      | 		#sleep(1.0)
      | 	#end
      | 	sleep(1.0)
      | 	#sleep(vibration_time)
      | 
      | 	movel(tilted_pose_in_base, a=0.03, v=0.1)
      | 	set_analog_out(0, 0.0)
      | 
      | 	tilt_pose_rel = pose_trans(pose_inv(p_center), tilted_pose_in_base)
      | 
      | 	lifted_pose_rel = pose_trans(lift_offset, tilt_pose_rel)
      | 
      | 	global lifted_pose = pose_trans(p_center, lifted_pose_rel)
      | 	movel(lifted_pose, a=0.03, v=0.1)
      | 	CCW_Rotate()
      | end
      | 
      | 
      | # calculate center pose on top of the container using pose transformation
      | def center_pose():
      | 	# pose transformation from side of the container to top to get center point
      | 	trans_rel = p[-0.005, 0.05, -0.027, 0, 0, 0]
      | 
      | 	p_translated = pose_trans(place_pose, trans_rel)
      | 	cx = p_translated[0]
      | 	cy = p_translated[1]
      | 	cz = p_translated[2]
      | 
      | 	global p_center_vertical = p[cx,cy,cz, 0, 0, 4.14]
      | 
      | 	#movej(p_center_vertical, a =0.3, v =0.3)
      | 	return p_center_vertical
      | end
      | 
      | # update center pose based on tilting
      | def updated_center_pose(p_center_vertical, angle_deg):
      | 	hinge_pose = pose_trans(p_center_vertical, p[0,0,-0.2,0,0,0])
      | 	local_rel = pose_trans(pose_inv(hinge_pose), p_center_vertical)
      | 
      | 	rot_tilt = p[0,0,0, -deg2rad(angle_deg),0,0]
      | 	local_rel_tilted = pose_trans(rot_tilt, local_rel)
      | 
      | 	global p_center = pose_trans(hinge_pose, local_rel_tilted)
      | 	return p_center
      | end
      | 
      | #------
      | # POTS commands
      | def tilt_send(angle):
      | 	socket_open("192.168.12.101", 80)
      | 	angle = 92.0 - angle
      | 	socket_send_string("Tilt,"+to_str(angle)+",0")
      | 	sync()
      | 	sleep(0.5)
      | 	socket_close()
      | end
      | 
      | def Motors_off():
      | 	socket_open("192.168.12.101", 80)
      | 	socket_send_string("Off,0,0")
      | 	sync()
      | 	sleep(0.5)
      | 	socket_close()
      | end
      | 
      | def Rotate():
      | 	socket_open("192.168.12.101", 80)
      | 	socket_send_string("FullRotation, 1, 2000")
      | 	sync()
      | 	sleep(0.5)
      | 	socket_close()
      | end
      | 
      | 
      | def CCW_Rotate():
      | 	socket_open("192.168.12.101", 80)
      | 	socket_send_string("FullRotation, -1, 2000")
      | 	sync()
      | 	sleep(0.5)
      | 	socket_close()
      | end
      | 
      | def tilt_to_home():
      | 	socket_open("192.168.12.101", 80)
      | 	socket_send_string("Home,0,0")
      | 	sync()
      | 	sleep(0.5)
      | 	socket_close()
      | end
    SuppressedNode
      Script file /programs/04 Scripts/dosing.script
        | def vibration_2():
        | 	set_analog_out(0,0.4)
        | 	sleep(0.8)
        | 	set_analog_out(0,0.0)
        | 	sleep(0.2)
        | end
        | 
        | def vibration_3():
        | 	set_analog_out(0,0.4)
        | 	sleep(0.5)
        | 	set_analog_out(0,0.0)
        | 	sleep(0.3)
        | end
        | 
        | def vibration_4():
        | 	set_analog_out(0,0.4)
        | 	sleep(0.6)
        | 	set_analog_out(0, 0.0)
        | 	sleep(0.5)
        | end
        | 
        | def vibration_1():
        | 	set_analog_out(0,0.4)
        | 	sleep(1)
        | 	set_analog_out(0,0.0)
        | 	sleep(0)
        | end
        | 
        | def move_tilt_in_steps(Pow_center, final_pose, steps):
        | 	i = 0
        | 	while i <= steps:
        | 		ratio = i / steps
        | 		pose_step = p[Pow_center[0] + ratio * (final_pose[0] - Pow_center[0]), Pow_center[1] + ratio * (final_pose[1] -Pow_center[1]),Pow_center[2] + ratio * (final_pose[2] - Pow_center[2]), Pow_center[3] + ratio * (final_pose[3] - Pow_center[3]), Pow_center[4] + ratio * (final_pose[4] - Pow_center[4]), Pow_center[5] + ratio * (final_pose[5] - Pow_center[5])]
        | 		movej(pose_step, a=1.2, v=0.15)
        | 		sleep(0.1)
        | 		i = i+1
        | 	end
        | end
        | 
        | def tilt_container(angle):
        | 	p_center = get_actual_tcp_pose()
        | 	hinge_offset = p[0,0,-0.23,0,0,0]
        | 	pivot_pose = pose_trans(p_center, hinge_offset)
        | 	pose_rel = pose_trans(pose_inv(pivot_pose), p_center)
        | 	angle_mid = (angle/2.0)*3.1416/180
        | 	angle_end = angle*3.1416/180
        | 	tilt_mid = p[0,0,0, -angle_mid, 0, 0]
        | 	tilt_end = p[0,0,0, -angle_end, 0, 0]
        | 	pose_rel_mid = pose_trans(tilt_mid, pose_rel)
        | 	pose_rel_end = pose_trans(tilt_end, pose_rel)
        | 	via_pose = pose_trans(pivot_pose, pose_rel_mid)
        | 	end_pose = pose_trans(pivot_pose, pose_rel_end)
        | 	movec(via_pose, end_pose, a=0.05, v=0.01, r=0.001)
        | 	p_center = get_actual_tcp_pose()
        | end
        | 
        | def deg2rad(d):
        | 	return d*3.141592/180
        | end
        | 
        | def map_tilt_to_ry_deg(container_deg):
        | 	#ry_deg = -0.875*container_deg +87.0
        | 	#return clamp(ry_deg, 5.0, 80.0)
        | 	if (Pow_name == "NaCl" or Pow_name == "Mannitol" or Pow_name == "CCS" or Pow_name == "MCC"):
        | 		if ( level>=10.0):
        | 			ry_min = 10.0
        | 			ry_max = 75.0
        | 		elif (level<10.00 and level >1.00):
        | 			ry_min = 16.0
        | 			ry_max = 65.0
        | 		else:
        | 			ry_min=17.0
        | 			ry_max=75.0
        | 		end
        | 	else:
        | 		if ( level>=10.0):
        | 			ry_min = 0.0
        | 			ry_max = 65.0
        | 		elif (level<10.00 and level >1.00):
        | 			ry_min = 10.0
        | 			ry_max = 45.0
        | 		else:
        | 			ry_min=0.0
        | 			ry_max=50.0
        | 		end
        | 
        | 	end
        | 	local span_count = angle_max -angle_min
        | 	local span_ry = ry_max - ry_min
        | 
        | 	local t = (container_deg -angle_min)/span_count
        | 	local ry_deg = ry_max - t*span_ry
        | 
        | 	return clamp(ry_deg, ry_min, ry_max)
        | 
        | end
        | 
        | def caluclate_corrections(level):
        | 	z_high = 0.01
        | 	z_low = -0.08
        | 	y_high = -0.01
        | 	y_low = -0.015
        | 
        | 	scale = (level - 10.0) / (100.0-10.0)
        | 
        | 	global correction_z = z_low + scale*(z_high - z_low)
        | 	global correction_y = y_low + scale*(y_high -y_low)
        | 
        | end
        | 
        | def scoop_powder(p_center):
        | 	#lift_offset = p[0, 0, 0.05, 0, 0, 0]
        | 	vibration_voltage = 0.4
        | 	vibration_time = 3.0
        | 	diameter = 0.07
        | 	global scoop_radius_default = 0.0
        | 	#p_center = center_pose_t
        | 
        | 
        | 	if (level >=70.00):
        | 		approach_offset = p[0.008,0,0.22,0,0,0]
        | 		lift_offset = p[0, 0, 0.05, 0, 0, 0]
        | 		caluclate_corrections(level)
        | 	elif (level >=10.00 and level <70):
        | 		approach_offset = p[0.008,0,0.22,0,0,0]
        | 		lift_offset = p[0, 0, 0.15, 0, 0, 0]
        | 		caluclate_corrections(level)
        | 	elif (level<10.00 and level >= 1.00):
        | 		approach_offset = p[0.01,0,0.22,0,0,0]
        | 		correction_z = -0.08
        | 		correction_y = -0.01
        | 		lift_offset = p[0, 0, 0.14, 0, 0, 0]
        | 	else:
        | 		approach_offset = p[0.008,0,0.22,0,0,0]
        | 		correction_z = -0.08
        | 		correction_y = -0.01
        | 		lift_offset = p[0, 0, 0.14, 0, 0, 0]
        |  	end
        | 
        | 	if (spatula == "spatula_L"):
        | 		global spatula_depth = 0.015
        | 	elif (spatula == "spatula_M"):
        | 		global spatula_depth = 0.01
        | 	elif (spatula == "spatula_S"):
        | 		global spatula_depth = 0.008
        | 	elif (spatula == "spatula_flat_M"):
        | 		global spatula_depth = 0.001
        | 	elif (spatula == "spatula_flat_S"):
        | 		global spatula_depth = 0.005
        | 	end
        | 
        | 	scoop_radius_default = diameter/2 - spatula_depth
        | 	scoop_entry_pose = pose_trans(p_center, approach_offset)
        | 	movel(scoop_entry_pose, a=0.1, v=0.25)
        | 
        | 	scoop_start_rel = p[scoop_radius_default, 0, scoop_depth, 0, 0, 0]
        | 
        | 	rot_mid = p[0, 0, 0, 0, 0, 0.785]
        | 	rot_end = p[0, 0, 0, 0, 0, 1.5708]
        | 
        | 	scoop_via_rel = pose_trans(rot_mid, scoop_start_rel)
        | 	scoop_end_rel = pose_trans(rot_end, scoop_start_rel)
        | 
        | 	scoop_start_pose = pose_trans(p_center, scoop_start_rel)
        | 	scoop_via_pose = pose_trans(p_center, scoop_via_rel)
        | 	scoop_end_pose = pose_trans(p_center, scoop_end_rel)
        | 
        | 	movel(scoop_start_pose, a=0.5, v=0.3)
        | 	#movel(p_center, a=0.5, v=1.0)
        | 	#sleep(5.0)
        | 
        | 	if (level<90.0):
        | 		Rotate()
        | 	end
        | 
        | 	#movec(scoop_via_pose, scoop_end_pose, a=0.03, v=0.05)
        | 	movec(scoop_via_pose, scoop_end_pose, a=0.03, v=0.02)
        | 	#movel(pose_trans(get_actual_tcp_pose(), p[0,0,0,0,0,deg2rad(90.0)]), a=0.03, v=0.05)
        | 	sleep(1.0)
        | 	local ry_deg = map_tilt_to_ry_deg(angle_deg)
        | 	local ry = deg2rad(ry_deg)
        | 	local end_rel = pose_trans(pose_inv(p_center), scoop_end_pose)
        | 	local end_rel_tilted = pose_trans(end_rel, p[0, 0, 0, 0, ry, 0])
        | 	global tilted_pose_in_base = pose_trans(p_center, p[0,correction_y,correction_z,end_rel_tilted[3],end_rel_tilted[4], end_rel_tilted[5]])
        | 	global tilted_pose_in_base = pose_trans(tilted_pose_in_base, p[0, 0, spatula_len, 0, 0, 0])
        | 
        | 	if (Pow_name == "lactose_fine" or Pow_name == "Magnesium_sterate"):
        | 		tilt_send((angle_deg+5))
        | 	end
        | 	movel(tilted_pose_in_base, a=0.03, v=0.1)
        | 
        | 	if (Pow_name == "lactose_fine" or Pow_name == "Magnesium_sterate"):
        | 		tilt_send((angle_deg-5))
        | 	end
        | 
        | 	if (spatula=="spatula_flat_S" or spatula=="spatula_S"):
        | 		vibration_3()
        | 	else:
        | 		set_analog_out(0, vibration_voltage)
        | 	end
        | 	if (Pow_name=="Mannitol" or Pow_name =="NaCl"):
        | 		local n=1.4
        | 	else:
        | 		local n=1.5
        | 	end
        | 	local ry_level = deg2rad(ry_deg/n)
        | 	local end_rel_tilted_level = pose_trans(end_rel, p[0, 0, 0, 0, ry_level, 0])
        | 	local level_tilted_pose_in_base = pose_trans(p_center, p[0,correction_y,correction_z,end_rel_tilted_level[3],end_rel_tilted_level[4], end_rel_tilted_level[5]])
        | 	local level_tilted_pose_in_base = pose_trans(level_tilted_pose_in_base, p[0, 0, spatula_len, 0, 0, 0])
        | 
        | 	movel(level_tilted_pose_in_base, a=0.03, v=0.1)
        | 	#if (level>70.0):
        | 		#sleep(1.0)
        | 	#end
        | 	sleep(1.0)
        | 	#sleep(vibration_time)
        | 
        | 	movel(tilted_pose_in_base, a=0.03, v=0.1)
        | 	set_analog_out(0, 0.0)
        | 
        | 	tilt_pose_rel = pose_trans(pose_inv(p_center), tilted_pose_in_base)
        | 
        | 	lifted_pose_rel = pose_trans(lift_offset, tilt_pose_rel)
        | 
        | 	global lifted_pose = pose_trans(p_center, lifted_pose_rel)
        | 	movel(lifted_pose, a=0.03, v=0.1)
        | 	CCW_Rotate()
        | end
        | 
        | 
        | def center_pose():
        | 	trans_rel = p[-0.005, 0.05, -0.015, 0, 0, 0]
        | 
        | 	p_translated = pose_trans(place_pose, trans_rel)
        | 	cx = p_translated[0]
        | 	cy = p_translated[1]
        | 	cz = p_translated[2]
        | 
        | 	global p_center_vertical = p[cx,cy,cz, 0, 0, 4.09]
        | 
        | 	#movej(p_center_vertical, a =0.3, v =0.3)
        | 	return p_center_vertical
        | end
        | 
        | def updated_center_pose(p_center_vertical, angle_deg):
        | 	hinge_pose = pose_trans(p_center_vertical, p[0,0,-0.2,0,0,0])
        | 	local_rel = pose_trans(pose_inv(hinge_pose), p_center_vertical)
        | 
        | 	rot_tilt = p[0,0,0, -deg2rad(angle_deg),0,0]
        | 	local_rel_tilted = pose_trans(rot_tilt, local_rel)
        | 
        | 	global p_center = pose_trans(hinge_pose, local_rel_tilted)
        | 	return p_center
        | end
        | 
        | def tilt_send(angle):
        | 	socket_open("192.168.12.101", 80)
        | 	angle = 92.0 - angle
        | 	socket_send_string("Tilt,"+to_str(angle)+",0")
        | 	sync()
        | 	sleep(0.5)
        | 	socket_close()
        | end
        | 
        | def Motors_off():
        | 	socket_open("192.168.12.101", 80)
        | 	socket_send_string("Off,0,0")
        | 	sync()
        | 	sleep(0.5)
        | 	socket_close()
        | end
        | 
        | def Rotate():
        | 	socket_open("192.168.12.101", 80)
        | 	socket_send_string("FullRotation, 1, 2000")
        | 	sync()
        | 	sleep(0.5)
        | 	socket_close()
        | end
        | 
        | 
        | def CCW_Rotate():
        | 	socket_open("192.168.12.101", 80)
        | 	socket_send_string("FullRotation, -1, 2000")
        | 	sync()
        | 	sleep(0.5)
        | 	socket_close()
        | end
        | def tilt_to_home():
        | 	socket_open("192.168.12.101", 80)
        | 	socket_send_string("Home,0,0")
        | 	sync()
        | 	sleep(0.5)
        | 	socket_close()
        | end
    Script file /programs/04 Scripts/Weight_scale_socket_s.script
      | def get_weight():
      | 	socket_open("192.168.12.111", 3002)
      | 	sleep(0.2)
      | 	textmsg("socket opened successfully!")
      | 	socket_send_string("GET_WEIGHT")
      | 	sync()
      | 	sleep(0.5)
      | 	receiveFromServ = socket_read_ascii_float(6)
      | 	while (receiveFromServ[0] <1):
      | 		sleep(0.5)
      | 		receiveFromServ = socket_read_ascii_float(1)
      | 		textmsg("retrying read:", receiveFromServ)
      | 	end
      | 	textmsg("Received weight:", receiveFromServ[1])
      | 	socket_close()
      | 	sleep(0.2)
      | 	return receiveFromServ[1]
      | end
      | 
      | def tare_scale():
      | 	socket_open("192.168.12.111", 3002)
      | 	socket_send_string("TARE")
      | 	sleep(0.5)
      | 	socket_close()
      | end
      | 
      | def zero_scale():
      | 	socket_open("192.168.12.111", 3002)
      | 	socket_send_string("ZERO")
      | 	sleep(0.5)
      | 	socket_close()
      | end
      | 
      | def log_weight():
      | 	socket_open("192.168.12.111", 3002)
      | 	socket_send_string("LOG_WEIGHT")
      | 	sleep(0.5)
      | 	socket_close()
      | end
      | 
      | def send_target_info():
      | 	socket_open("192.168.12.111", 3002)
      | 	socket_send_string("SET_TARGET:" + to_str(target_weight))
      | 	sleep(0.2)
      | 	socket_close()
      | end
      | def send_powder_info():
      | 	socket_open("192.168.12.111", 3002)
      | 	socket_send_string("SET_POWDER:" + Pow_name)
      | 	sleep(0.2)
      | 	socket_close()
      | end
      | def send_spatula_info():
      | 	socket_open("192.168.12.111", 3002)
      | 	socket_send_string("SET_SPATULA:" + spatula)
      | 	sleep(0.2)
      | 	socket_close()
      | end
      | 
      | def send_level_info():
      | 	socket_open("192.168.12.111",3002)
      | 	socket_send_string("SET_LEVEL:" + to_str(level))
      | 	sleep(0.2)
      | 	socket_close()
      | end
    SuppressedNode
      Script file /programs/04 Scripts/Calibration_s.script
        | # ------------------------------------------------------------
        | # Theoretical W_FULL from Cylinder Volume + Density
        | # (Eliminates manual W_FULL; keeps W_EMPTY + W_now for level)
        | # ------------------------------------------------------------
        | # -------------------------
        | # 1) Define container geometry (cylindrical inner dimensions)
        | # -------------------------
        | # Use mm for readability; we convert internally.
        | global D_INNER_MM   = 66.0     # inner diameter of container (mm)
        | global H_FILL_MM    = 125.0    # usable fill height up to "full" (mm)
        | 
        | # -------------------------
        | # 2) Define powder density
        | # -------------------------
        | # Density is directly set for now (as per your requirement).
        | # Use g/mL (common lab bulk density style).
        | #global RHO_G_PER_ML = 0.40     # example: 0.55 g/mL (replace per powder)
        | 
        | # ------------------------------------------------------------
        | # Spatula volumes (manufacturer specified)
        | # ------------------------------------------------------------
        | 
        | # Large spatula
        | global SPATULA_L_VOL_ML = 5.0        # 1 teaspoon = 5 mL
        | 
        | # Medium spatula
        | global SPATULA_M_VOL_ML = 1.25       # 1/4 teaspoon = 1.25 mL
        | 
        | # Small spatula
        | global SPATULA_S_VOL_ML = 0.15625    # 1/32 teaspoon = 0.15625 mL
        | 
        | global SPATULA_FLAT_M_VOL_ML  = 2.2
        | global SPATULA_FLAT_S_VOL_ML  = 1.2   #based on caluclations using rho = m/V
        | 
        | # -------------------------
        | # 4) Utility functions
        | # -------------------------
        | 
        | 
        | def cyl_volume_mL(d_mm, h_mm):
        |   # Converts mm -> m, computes cylinder volume in m^3, converts to mL
        |   # V = π * r^2 * h
        |   local d_m  = d_mm / 1000.0
        |   local h_m  = h_mm / 1000.0
        |   local r_m  = d_m / 2.0
        |   local v_m3 = 3.141592653589793 * r_m * r_m * h_m
        |   global v_mL = v_m3 * 1000000.0     # 1 m^3 = 1,000,000 mL
        |   return v_mL
        | end
        | 
        | def compute_W_full_theoretical():
        |   V_mL = cyl_volume_mL(D_INNER_MM, H_FILL_MM)
        |   local M_powder_g = density * V_mL
        |   global W_FULL = W_EMPTY + M_powder_g
        |   return W_FULL
        | end
        | 
        | 
        | # ------------------------------------------------------------
        | # Function: Theoretical scoop weight from volume
        | # ------------------------------------------------------------
        | def scoop_weight_from_volume(vol_mL, density):
        |   return vol_mL * density
        | end
        | 
        | # ------------------------------------------------------------
        | # Function: Get scoop weight based on spatula type
        | # ------------------------------------------------------------
        | def get_scoop_weight(spatula):
        |   local vol = 0.0
        | 
        |   if (spatula == "spatula_L"):
        |     vol = SPATULA_L_VOL_ML
        |   elif (spatula == "spatula_M"):
        |     vol = SPATULA_M_VOL_ML
        |   elif (spatula == "spatula_S"):
        |     vol = SPATULA_S_VOL_ML
        |   elif (spatula == "spatula_flat_M"):
        |     return SPATULA_FLAT_M_VOL_ML
        |   elif (spatula == "spatula_flat_S"):
        |     return SPATULA_FLAT_S_VOL_ML
        |   else:
        |     textmsg("Unknown spatula type")
        |     return 0.0
        |   end
        | 
        |   global target_g =  scoop_weight_from_volume(vol, density)
        |   return target_g
        | end
    Script file /programs/04 Scripts/Read_QR.script
      | global SERVER_IP   = "192.168.12.111"
      | global SERVER_PORT = 3002
      | 
      | global qr_container_id = 0
      | global qr_chemical_id  = 0
      | global qr_H_mm         = 0
      | global qr_H_c_mm         = 0
      | global qr_neck_d_mm    = 0
      | global qr_neck_sh_mm   = 0
      | global qr_length_mm    = 0
      | global qr_diameter_mm  = 0
      | global qr_empty_weight_g  = 0
      | global qr_volume_ml    = 0
      | global qr_shape_code   = 0
      | global shape = ""
      | global cent_edge = 0
      | global pick_2_base = 0.27375 # distance from tcp to base of picking table
      | global place_2_counter = 0.18775 # distance from base of holders on robot platform  to TCP
      | 
      | def read_qr_db_data():
      | 
      |   socket_open(SERVER_IP, SERVER_PORT)
      |   sleep(0.5)
      |   socket_send_string("GET_QR_FLOATS")
      |   sleep(5)
      | 
      |   local fl = socket_read_ascii_float(11)
      |   socket_close()
      | 
      |   global qr_container_id = fl[1]
      |   global qr_chemical_id = fl[2]
      |   global qr_H_mm         = fl[3]/1000
      |   global qr_H_c_mm         = fl[4]/1000
      |   global qr_neck_d_mm    = fl[5]/1000
      |   global qr_neck_sh_mm   = fl[6]/1000
      |   global qr_length_mm    = fl[7]/1000
      |   global qr_diameter_mm  = fl[8]/1000
      |   global qr_empty_weight_g = fl[9]
      |   global qr_volume_ml    = fl[10]
      |   global qr_shape_code   = fl[11]
      | 
      |   if (qr_shape_code == 1.0):
      | 	shape = "cylindrical"
      | 	cent_edge = qr_diameter_mm
      |   else:
      | 	shape = "cubical"
      | 	cent_edge = qr_length_mm
      |   end
      | 
      |   textmsg("container_id = ", qr_container_id)
      |   textmsg("chemical_id = ", qr_chemical_id)
      |   textmsg("h_mm = ", qr_H_mm)
      |   textmsg("H_c_mm = ", qr_H_c_mm)
      |   textmsg("neck_d_mm = ", qr_neck_d_mm)
      |   textmsg("neck_sh_mm = ", qr_neck_sh_mm)
      |   textmsg("length_mm = ", qr_length_mm)
      |   textmsg("diameter_mm = ", qr_diameter_mm)
      |   textmsg("empty_weight_g = ", qr_empty_weight_g)
      |   textmsg("volume_ml = ", qr_volume_ml)
      |   textmsg("shape_code = ", qr_shape_code)
      | end
  Folder BeforeStarts [hidden by the author, left out]
  Folder powder dispensing variable init
    Start_thread := False
    vib_thread := False
    Folder QR assignment init
      d_cc := 0.06
      W_EMPTY := 50.131
    kp := 0.0015
    ki := 0.0001
    kd := 0.01
    dt := 0.03
    Integral_error := 0
    current_error := 0
    previous_error := 0
    tilt_increment := 0
    tilt_angle := 0
    diff := 0
    current_pose := get_actual_tcp_pose()
    Relative_trans := p[0, 0, -0.035, 0, 0, 0]
    SuppressedNode
      ContA_plc_offst := p[-0.00205, 0.02547, 0.03730, -0.03, -2.183, 6.165]
    SuppressedNode
      PowA_50_offset := p[0.21808, -0.19943, 0.06584, 0, 0, 0]
    SuppressedNode
      Script: scooping_init()
    Script: tilt_init_reference()
    switch_spat_M := True
    switch_spat_S := True
    switch_spat_F_M := True
    switch_spat_F_S := True
    last_scale := 0
Robot Program (runOnlyOnce=false)
  Folder MAIN [hidden by the author, left out]
Thread Thread_1 (runOnlyOnce=false)
  If Start_thread≟ True
    weight_value := get_weight()
    Wait Sleep waitTime=0.1
    Script: sync()
  Script: sync()
Thread Thread_2 (runOnlyOnce=false)
  Loop While (checkContinuously=true) expression=vib_thread≟ True
    diff := target_weight-weight_value
    If diff>0.02 and spatula≠"spatula_flat_S" (checkContinuously=true)
      SuppressedNode
        Script: vibration_1()
      Set AnalogOutput pin=analog_out[0]; analogValue=4
    ElseIf diff>0.02 and spatula≟"spatula_flat_S"
      Script: vibration_3()
    ElseIf diff≤0.03 (checkContinuously=true)
      Script: vibration_2()
    SuppressedNode
      ElseIf diff≥0.01 and diff<0.05
        Script: vibration_3()
    SuppressedNode
      ElseIf diff>0 and diff<0.01
        Script: vibration_4()
    Else 
      Set AnalogOutput pin=analog_out[0]; analogValue=0
  Script: sync()
SubProgram -> Sub_Vision_V18
SubProgram  [hidden by the author, left out]
SubProgram -> Sub_Action_V4
